(* IEC 61131-3 sources: plc-vscode/tests/st/all/trust-platform/examples/siemens_scl_v1/src, 2 files *)

(* ---- Main.st ---- *)
FUNCTION_BLOCK FB_EdgeCounter
VAR_INPUT
    Enable : BOOL;
END_VAR
VAR_OUTPUT
    Count : DINT;
END_VAR
VAR
    LastEnable : BOOL;
END_VAR

IF #Enable AND NOT #LastEnable THEN
    #Count := #Count + 1;
END_IF;
#LastEnable := #Enable;
END_FUNCTION_BLOCK

PROGRAM Main
VAR
    Counter : FB_EdgeCounter;
    Total : DINT;
    Pulse : BOOL;
    CountNonZero : BOOL;
END_VAR

#Counter(Enable := #Pulse);
#Total := #Counter.Count;
#CountNonZero := #Total > 0;
END_PROGRAM

(* ---- Configuration.st ---- *)
CONFIGURATION SiemensDemo
RESOURCE SiemensRes ON PLC
TASK Cycle (INTERVAL := T#50ms, PRIORITY := 1);
PROGRAM P1 WITH Cycle : Main;
END_RESOURCE
VAR_CONFIG
    P1.Pulse AT %IX0.0 : BOOL;
    P1.CountNonZero AT %QX0.0 : BOOL;
END_VAR
END_CONFIGURATION
